Fanuc KAREL source: KT00772.KL

PROGRAM KT00772
%NOLOCKGROUP
VAR
  I1: INTEGER
  I2: INTEGER
  OUT: INTEGER
BEGIN
  I1 = 2
  I2 = 3
  I1 = 2
  I2 = 3
  OUT = ASIN(I1)
END KT00772
